FUNCTION_BLOCK CU_TEST
VAR_INPUT
  P : BOOL;
  RS : BOOL;
END_VAR
VAR
  c : CTU;
END_VAR
BEGIN
  c(CU := P, R := RS, PV := 2);
  //#ASSERT NOT c.Q : Pbad
END_FUNCTION_BLOCK
